Fanuc KAREL source: KB00006.KL

PROGRAM KB00006
%NOLOCKGROUP
%ENVIRONMENT PBQMGR
VAR
  P1: INTEGER
  P2: QUEUE_TYPE
  P3: ARRAY[4] OF INTEGER
  P4: INTEGER
  P5: INTEGER
BEGIN
  P1 = 1
  P3[1] = 1
  P4 = 1
  P5 = 1
  APPEND_QUEUE(P1, P2, P3, P4, P5)
END KB00006
